ABB RAPID module: MainCall.mod

%%%
  VERSION:1
  LANGUAGE:ENGLISH
%%%
MODULE MOD_MainCall

    ! -------------------------------
    ! Define customized variables here
    ! ...

	! Tool variables:

	! Reference variables:
	PERS wobjdata FrameS := [FALSE, TRUE, "", [[0,0,0],[1,0,0,0]],[[1234.570,-98.765,50.500],[0.96592583,0.00000000,0.00000000,0.25881905]]];

	PROC SubProg2()
		ConfJ \On;
		ConfL \Off;
		MoveAbsJ [[20.000000,-10.000000,20.000000,0.000000,30.000000,0.000000],[9E+09,9E+09,9E+09,9E+09,9E+09,9E+09]],v500,z1,tool0 \WObj:=FrameS;
	ENDPROC

	PROC Main()
		ConfJ \On;
		ConfL \Off;
		! Program generated by RoboDK v6.0.7 for ABB IRB 120-3/0.6 on XX/XX/XXXX 12:58:43
		! Using nominal kinematics.
		MoveAbsJ [[0.000000,-10.000000,20.000000,0.000000,30.000000,0.000000],[9E+09,9E+09,9E+09,9E+09,9E+09,9E+09]],v500,z1,tool0 \WObj:=FrameS;
		SubProg2;
		NotAProgram;
	ENDPROC

ENDMODULE
